Fanuc KAREL source: compact_preamble.KL

PROGRAM KB00135
%NOLOCKGROUP
VAR
P1:INTEGER;P2 : STRING[80];P3:INTEGER;P4:INTEGER
BEGIN
P1=1
P2='A'
P3=1
P4=1
POST_ERR_L(P1,P2,P3,P4)
END KB00135
